SUBAPPLICATION SlurryTanker (* Subapplication Type *)
  (* Standard: 61499-2 *)
  (* Version 1.0, 2023-02-11, franz *)
  IMPORT logiBUS::io::DQ::logiBUS_DO::Output_Q2;
  IMPORT logiBUS::io::DQ::logiBUS_DO::Output_Q3;
  IMPORT logiBUS::io::DQ::logiBUS_DO::Output_Q4;
  IMPORT logiBUS::io::DQ::logiBUS_DO::Output_Q5;
  IMPORT logiBUS::io::DQ::logiBUS_DO::Output_Q6;
  IMPORT logiBUS::io::DQ::logiBUS_DO::Output_Q7;
  IMPORT logiBUS::io::DQ::logiBUS_DO::Output_Q9;
  IMPORT logiBUS::io::DQ::logiBUS_DO::Output_Q10;
  IMPORT logiBUS::io::DQ::logiBUS_DO::Output_Q11;
  IMPORT logiBUS::io::DQ::logiBUS_DO::Invalid;
  IMPORT BlinkMarine::io::DI::PKP_2200_LI_DI::DigitalInput_Key_1;
  IMPORT BlinkMarine::io::DI::PKP_2200_LI_DI::DigitalInput_Key_2;
  IMPORT BlinkMarine::io::DI::PKP_2200_LI_DI::DigitalInput_Key_3;
  IMPORT BlinkMarine::io::DI::PKP_2200_LI_DI::DigitalInput_Key_4;
  IMPORT DefaultPool::AuxInput_Abscheider;
  IMPORT DefaultPool::AuxInput_Auseinanderklappen;
  IMPORT DefaultPool::AuxInput_Dom;
  IMPORT DefaultPool::AuxInput_Heckschieber;
  IMPORT DefaultPool::AuxInput_Knickdeichsel_heben;
  IMPORT DefaultPool::AuxInput_Knickdeichsel_senken;
  IMPORT DefaultPool::AuxInput_Licht;
  IMPORT DefaultPool::AuxInput_Schneidwerk;
  IMPORT DefaultPool::AuxInput_Seitenschieber;
  IMPORT DefaultPool::AuxInput_Verteiler_heben;
  IMPORT DefaultPool::AuxInput_Verteiler_senken;
  IMPORT DefaultPool::AuxInput_Zusammenklappen;
  IMPORT DefaultPool::SoftKey_Abscheider;
  IMPORT DefaultPool::SoftKey_Auseinanderklappen;
  IMPORT DefaultPool::SoftKey_Dom;
  IMPORT DefaultPool::SoftKey_Heckschieber;
  IMPORT DefaultPool::SoftKey_Knickdeichsel_heben;
  IMPORT DefaultPool::SoftKey_Knickdeichsel_senken;
  IMPORT DefaultPool::SoftKey_Licht;
  IMPORT DefaultPool::SoftKey_Schneidwerk;
  IMPORT DefaultPool::SoftKey_Seitenschieber;
  IMPORT DefaultPool::SoftKey_Verteiler_heben;
  IMPORT DefaultPool::SoftKey_Verteiler_senken;
  IMPORT DefaultPool::SoftKey_Zusammenklappen;
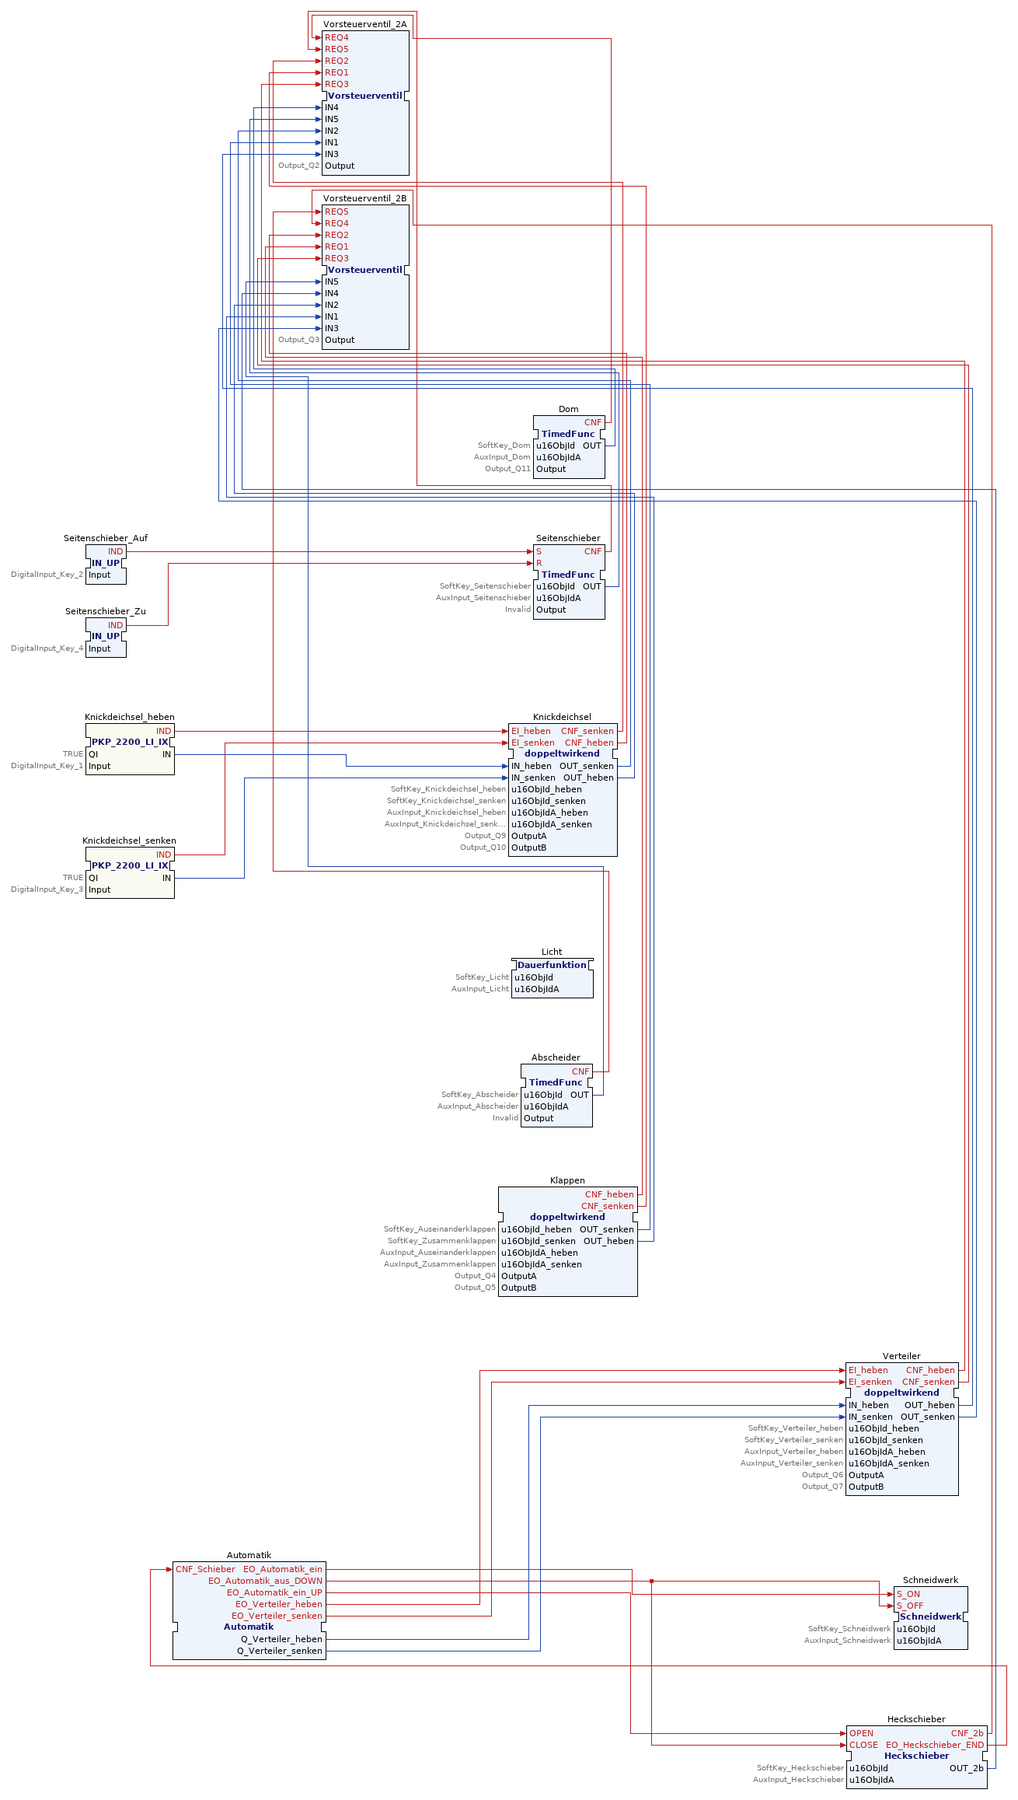
  (* Group funktionen: *)
  (* Group Vorsteuerventile: Vorsteuerventile *)
  (* Group Vorgewendeautomatik: Vorgewendeautomatik *)
  FBS
    Knickdeichsel_heben : BlinkMarine::io::DI::PKP_2200_LI_IX(QI := TRUE, Input := DigitalInput_Key_1); {SET_ATTRIBUTE(GroupName, funktionen)}
    Knickdeichsel_senken : BlinkMarine::io::DI::PKP_2200_LI_IX(QI := TRUE, Input := DigitalInput_Key_3); {SET_ATTRIBUTE(GroupName, funktionen)}
  END_FBS
  SUBAPPS
    Automatik : Automatik; {SET_ATTRIBUTE(GroupName, Vorgewendeautomatik)}
    Dom : TimedFunc(u16ObjId := SoftKey_Dom, u16ObjIdA := AuxInput_Dom, Output := Output_Q11); {SET_ATTRIBUTE(GroupName, funktionen)}
    Seitenschieber : TimedFunc(u16ObjId := SoftKey_Seitenschieber, u16ObjIdA := AuxInput_Seitenschieber, Output := Invalid); {SET_ATTRIBUTE(GroupName, funktionen)}
    Klappen : doppeltwirkend(u16ObjId_heben := SoftKey_Auseinanderklappen, u16ObjId_senken := SoftKey_Zusammenklappen, u16ObjIdA_heben := AuxInput_Auseinanderklappen, u16ObjIdA_senken := AuxInput_Zusammenklappen, OutputA := Output_Q4, OutputB := Output_Q5); {SET_ATTRIBUTE(GroupName, funktionen)}
    Verteiler : doppeltwirkend(u16ObjId_heben := SoftKey_Verteiler_heben, u16ObjId_senken := SoftKey_Verteiler_senken, u16ObjIdA_heben := AuxInput_Verteiler_heben, u16ObjIdA_senken := AuxInput_Verteiler_senken, OutputA := Output_Q6, OutputB := Output_Q7); {SET_ATTRIBUTE(GroupName, Vorgewendeautomatik)}
    Vorsteuerventil_2A : Vorsteuerventil(Output := Output_Q2); {SET_ATTRIBUTE(GroupName, Vorsteuerventile)}
    Vorsteuerventil_2B : Vorsteuerventil(Output := Output_Q3); {SET_ATTRIBUTE(GroupName, Vorsteuerventile)}
    Knickdeichsel : doppeltwirkend(u16ObjId_heben := SoftKey_Knickdeichsel_heben, u16ObjId_senken := SoftKey_Knickdeichsel_senken, u16ObjIdA_heben := AuxInput_Knickdeichsel_heben, u16ObjIdA_senken := AuxInput_Knickdeichsel_senken, OutputA := Output_Q9, OutputB := Output_Q10); {SET_ATTRIBUTE(GroupName, funktionen)}
    Licht : Dauerfunktion(u16ObjId := SoftKey_Licht, u16ObjIdA := AuxInput_Licht); {SET_ATTRIBUTE(GroupName, funktionen)}
    Abscheider : TimedFunc(u16ObjId := SoftKey_Abscheider, u16ObjIdA := AuxInput_Abscheider, Output := Invalid); {SET_ATTRIBUTE(GroupName, funktionen)}
    Schneidwerk : Schneidwerk(u16ObjId := SoftKey_Schneidwerk, u16ObjIdA := AuxInput_Schneidwerk); {SET_ATTRIBUTE(GroupName, Vorgewendeautomatik)}
    Heckschieber : Heckschieber(u16ObjId := SoftKey_Heckschieber, u16ObjIdA := AuxInput_Heckschieber); {SET_ATTRIBUTE(GroupName, Vorgewendeautomatik)}
    Seitenschieber_Auf : IN_UP(Input := DigitalInput_Key_2); {SET_ATTRIBUTE(GroupName, funktionen)}
    Seitenschieber_Zu : IN_UP(Input := DigitalInput_Key_4); {SET_ATTRIBUTE(GroupName, funktionen)}
  END_SUBAPPS
  EVENT_CONNECTIONS
    Dom.CNF TO Vorsteuerventil_2A.REQ4;
    Seitenschieber.CNF TO Vorsteuerventil_2A.REQ5;
    Abscheider.CNF TO Vorsteuerventil_2B.REQ5;
    Automatik.EO_Automatik_ein TO Schneidwerk.S_ON;
    Automatik.EO_Automatik_aus_DOWN TO Schneidwerk.S_OFF;
    Automatik.EO_Automatik_ein_UP TO Heckschieber.OPEN;
    Automatik.EO_Automatik_aus_DOWN TO Heckschieber.CLOSE;
    Heckschieber.CNF_2b TO Vorsteuerventil_2B.REQ4;
    Heckschieber.EO_Heckschieber_END TO Automatik.CNF_Schieber;
    Automatik.EO_Verteiler_heben TO Verteiler.EI_heben;
    Automatik.EO_Verteiler_senken TO Verteiler.EI_senken;
    Knickdeichsel_heben.IND TO Knickdeichsel.EI_heben;
    Knickdeichsel_senken.IND TO Knickdeichsel.EI_senken;
    Knickdeichsel.CNF_senken TO Vorsteuerventil_2A.REQ2;
    Knickdeichsel.CNF_heben TO Vorsteuerventil_2B.REQ2;
    Klappen.CNF_heben TO Vorsteuerventil_2B.REQ1;
    Klappen.CNF_senken TO Vorsteuerventil_2A.REQ1;
    Verteiler.CNF_heben TO Vorsteuerventil_2A.REQ3;
    Verteiler.CNF_senken TO Vorsteuerventil_2B.REQ3;
    Seitenschieber_Auf.IND TO Seitenschieber.S;
    Seitenschieber_Zu.IND TO Seitenschieber.R;
  END_CONNECTIONS
  DATA_CONNECTIONS
    Dom.OUT TO Vorsteuerventil_2A.IN4;
    Seitenschieber.OUT TO Vorsteuerventil_2A.IN5;
    Abscheider.OUT TO Vorsteuerventil_2B.IN5;
    Heckschieber.OUT_2b TO Vorsteuerventil_2B.IN4;
    Automatik.Q_Verteiler_heben TO Verteiler.IN_heben;
    Automatik.Q_Verteiler_senken TO Verteiler.IN_senken;
    Knickdeichsel_heben.IN TO Knickdeichsel.IN_heben;
    Knickdeichsel_senken.IN TO Knickdeichsel.IN_senken;
    Knickdeichsel.OUT_senken TO Vorsteuerventil_2A.IN2;
    Knickdeichsel.OUT_heben TO Vorsteuerventil_2B.IN2;
    Klappen.OUT_senken TO Vorsteuerventil_2A.IN1;
    Klappen.OUT_heben TO Vorsteuerventil_2B.IN1;
    Verteiler.OUT_heben TO Vorsteuerventil_2A.IN3;
    Verteiler.OUT_senken TO Vorsteuerventil_2B.IN3;
  END_CONNECTIONS
END_SUBAPPLICATION
